(* Logix 5000 project; controller TFF vendor 1 type 14 code 107 rev 34.11; software revision 34.03; part 26 of 36 *)
(* tags used below, declared in another part *)
   Address : DINT;   // Temp Address
   Index : DINT;   // Index
   AI101 : ALIAS FOR AnalogPoint[10];   // Filtrate Conductivity
   AI102 : ALIAS FOR AnalogPoint[11];   // Filtrate UV
   AI103 : ALIAS FOR AnalogPoint[12];   // Filtrate UV
   AI104 : ALIAS FOR AnalogPoint[9];   // Filtrate pH
   AlarmControl : AlarmControl;   // Alarm Control
   CPU_Scanning : BOOL;   // System Scanning Flag
   DigitalOutput : BOOL[256];   // Digital Output Array these bits are sent to output cards.
   DigitalPoint : DigitalPoint[150];   // Digital Point Array
   Drive : Drive[11];   // Drives Array
   FI101 : ALIAS FOR AnalogPoint[2];   // Filtrate Flow
   MIX001 : ALIAS FOR AnalogPoint[14];   // Mixer Speed
   Mixer : Mixer;   // Mixer config. structure
   Options : Options;   // Options List
   Phase0 : ALIAS FOR Phase[0];   // Phase 0
   PI001 : ALIAS FOR AnalogPoint[5];   // Feed Pressure
   PI002 : ALIAS FOR AnalogPoint[6];   // Retentate Pressure
   PI101 : ALIAS FOR AnalogPoint[7];   // Filtrate Pressure
   PI401 : ALIAS FOR AnalogPoint[8];   // Transfer Pump Pressure
   PLCFault : FaultRecordType;   // PLC Major Fault Record
   Rack_Murr_Node1_TF2S : IO_Station;   // Status of Node 1 TF2S
   Rack_Murr_Node1_TF3S : IO_Station;   // Status of Node 1 TF3S
   Rack_Murr_Node4_Instrum_TFF1 : IO_Station;   // Status of Node 4 Instrum TFF1
   Rack_Murr_Node4_Instrum_TFF2 : IO_Station;   // Status of Node 4 Instrum TFF2
   Rack_Murr_Node4_Instrum_TFF3 : IO_Station;   // Status of Node 4 Instrum TFF3
   Rack_Murr_Node4_Instrum_TFF4 : IO_Station;   // Status of Node 4 Instrum TFF4
   Rack_Murr_Node4_Instrum_TFF5 : IO_Station;   // Status of Node 4 Instrum TFF5
   Rack_Murr_Node5_Tank100 : IO_Station;   // Status of Node 5 Tank 100L
   Rack_Murr_Node5_Tank250 : IO_Station;   // Status of Node 5 Tank 250L
   Rack_Murr_Node5_Tank50 : IO_Station;   // Status of Node 5 Tank 50L
   RawAnalogInputArray : INT[50];   // Array of analog input raw
   SIC003 : ALIAS FOR Drive[3];   // Mixer
   SIC003DF : ALIAS FOR DigitalPoint[14];   // Mixer Defect
   SRL001 : ALIAS FOR DigitalPoint[15];   // Tank Skid Remote / Standalone
   SysControl : SysControl;   // General system status and command
   Tank : TankManagement;   // Tank Management
   ThisSystem : SystemType;
   TI001 : ALIAS FOR AnalogPoint[13];   // Feed Bag Temperature
   WI001 : ALIAS FOR AnalogPoint[15];   // Feed Bag Weight
   YA10 : ALIAS FOR DigitalPoint[59];   // PLC Program Major Fault
(* Process, continued *)

ROUTINE Drive_SIC003_Mixer   (* ladder *)
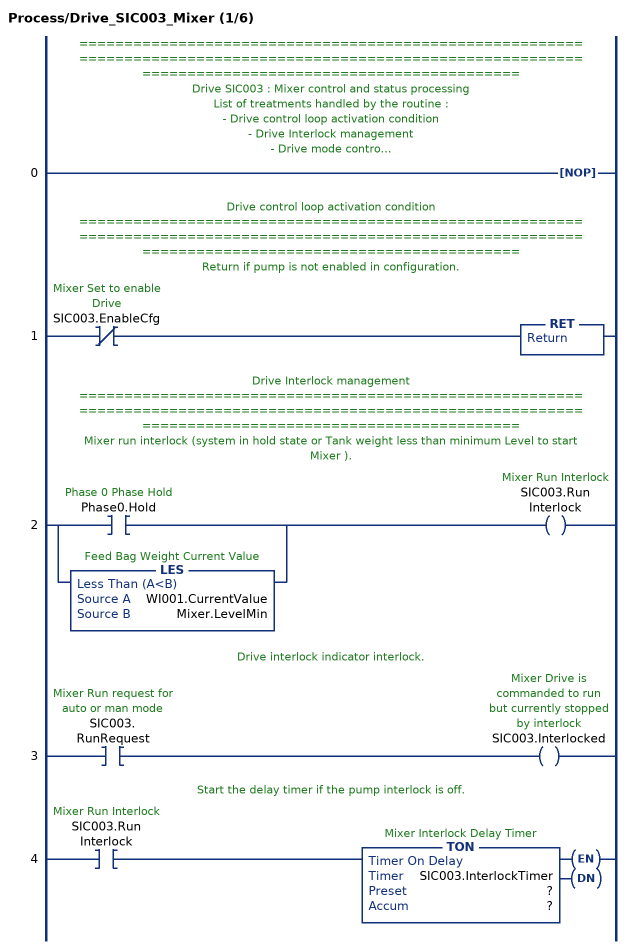
   // ==========================================================================================================================================================
   //                                                        Drive SIC003 : Mixer control and status processing
   //                                                     List of treatments handled by the routine :
   //                                                          - Drive control loop activation condition
   //                                                          - Drive Interlock management
   //                                                          - Drive mode control
   //                                                          - Drive run command control
   //                                                          - Drive status management
   //                                                          - Drive status for HMI
   //                                                          - Drive DigitalOutput control
   //                                                     -----------------------------------------------------------------------------------------------------------------------------------------------------
   //                                                     History
   //                                                          2019-AUG-13 - Actemium - B. Roch - Initial version for Candidate Release 3.00.00.00.a
   //                                                          2019-OCT-25 - Actemium - B. Roch - Modification for Candidate Release 3.00.00.00.d
   //                                                      - Add Mixer standalone condition to stop mixer
   // ==========================================================================================================================================================
   0: NOP();
   // Drive control loop activation condition
   // ==========================================================================================================================================================
   // Return if pump is not enabled in configuration.
   1: XIO(SIC003.EnableCfg)RET();
   // Drive Interlock management
   // ==========================================================================================================================================================
   // Mixer run interlock (system in hold state or Tank weight less than minimum Level to start Mixer ).
   2: [XIC(Phase0.Hold) ,LES(WI001.CurrentValue,Mixer.LevelMin) ]OTE(SIC003.RunInterlock);
   // Drive interlock indicator interlock.
   3: XIC(SIC003.RunRequest)OTE(SIC003.Interlocked);
   // Start the delay timer if the pump interlock is off.
   4: XIC(SIC003.RunInterlock)TON(SIC003.InterlockTimer,?,?);
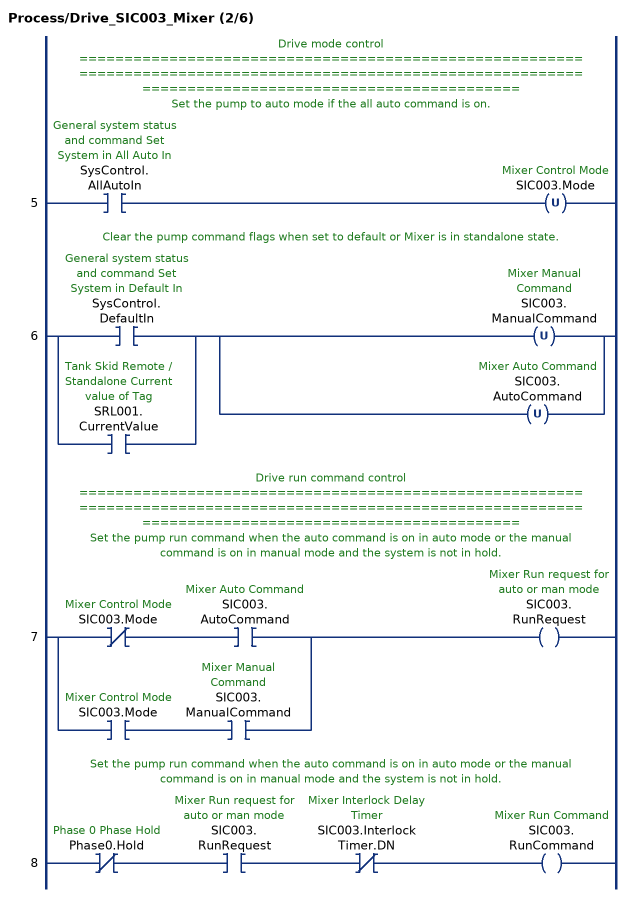
   // Drive mode control
   // ==========================================================================================================================================================
   // Set the pump to auto mode if the all auto command is on.
   5: XIC(SysControl.AllAutoIn)OTU(SIC003.Mode);
   // Clear the pump command flags when set to default or Mixer is in standalone state.
   6: [XIC(SysControl.DefaultIn) ,XIC(SRL001.CurrentValue) ][OTU(SIC003.ManualCommand) ,OTU(SIC003.AutoCommand) ];
   // Drive run command control
   // ==========================================================================================================================================================
   // Set the pump run command when the auto command is on in auto mode or the manual command is on in manual mode and the system is not in hold.
   7: [XIO(SIC003.Mode) XIC(SIC003.AutoCommand) ,XIC(SIC003.Mode) XIC(SIC003.ManualCommand) ]OTE(SIC003.RunRequest);
   // Set the pump run command when the auto command is on in auto mode or the manual command is on in manual mode and the system is not in hold.
   8: XIO(Phase0.Hold)XIC(SIC003.RunRequest)XIO(SIC003.InterlockTimer.DN)OTE(SIC003.RunCommand);
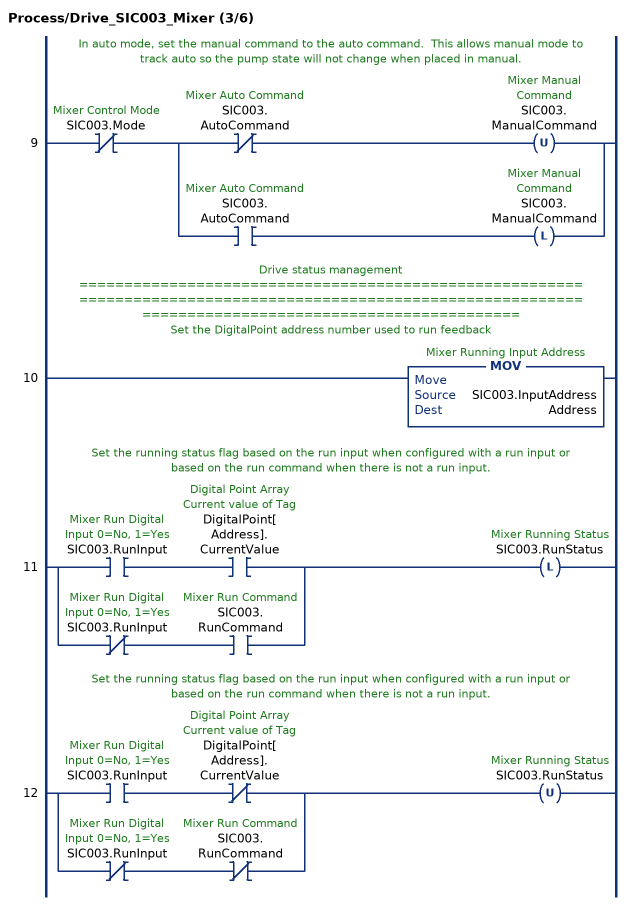
   // In auto mode, set the manual command to the auto command.  This allows manual mode to track auto so the pump state will not change when placed in manual.
   9: XIO(SIC003.Mode)[XIO(SIC003.AutoCommand) OTU(SIC003.ManualCommand) ,XIC(SIC003.AutoCommand) OTL(SIC003.ManualCommand) ];
   // Drive status management
   // ==========================================================================================================================================================
   // Set the DigitalPoint address number used to run feedback
   10: MOV(SIC003.InputAddress,Address);
   // Set the running status flag based on the run input when configured with a run input or based on the run command when there is not a run input.
   11: [XIC(SIC003.RunInput) XIC(DigitalPoint[Address].CurrentValue) ,XIO(SIC003.RunInput) XIC(SIC003.RunCommand) ]OTL(SIC003.RunStatus);
   // Set the running status flag based on the run input when configured with a run input or based on the run command when there is not a run input.
   12: [XIC(SIC003.RunInput) XIO(DigitalPoint[Address].CurrentValue) ,XIO(SIC003.RunInput) XIO(SIC003.RunCommand) ]OTU(SIC003.RunStatus);
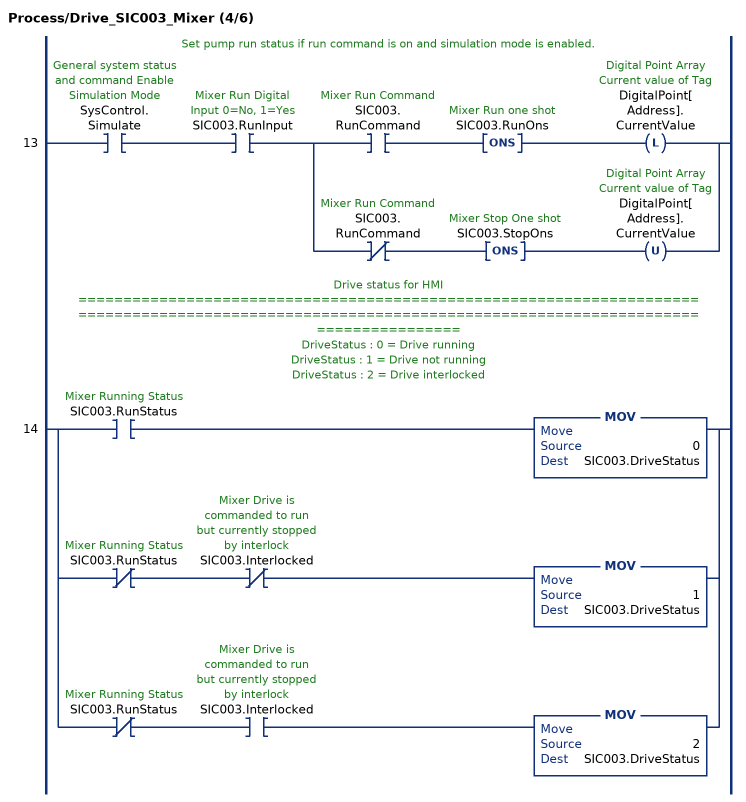
   // Set pump run status if run command is on and simulation mode is enabled.
   13: XIC(SysControl.Simulate)XIC(SIC003.RunInput)[XIC(SIC003.RunCommand) ONS(SIC003.RunOns) OTL(DigitalPoint[Address].CurrentValue) ,XIO(SIC003.RunCommand) ONS(SIC003.StopOns) OTU(DigitalPoint[Address].CurrentValue) ];
   // Drive status for HMI
   // ==========================================================================================================================================================
   //  DriveStatus : 0 = Drive running
   //  DriveStatus : 1 = Drive not running
   //  DriveStatus : 2 = Drive interlocked
   14: [XIC(SIC003.RunStatus) MOV(0,SIC003.DriveStatus) ,XIO(SIC003.RunStatus) XIO(SIC003.Interlocked) MOV(1,SIC003.DriveStatus) ,XIO(SIC003.RunStatus) XIC(SIC003.Interlocked) MOV(2,SIC003.DriveStatus) ];
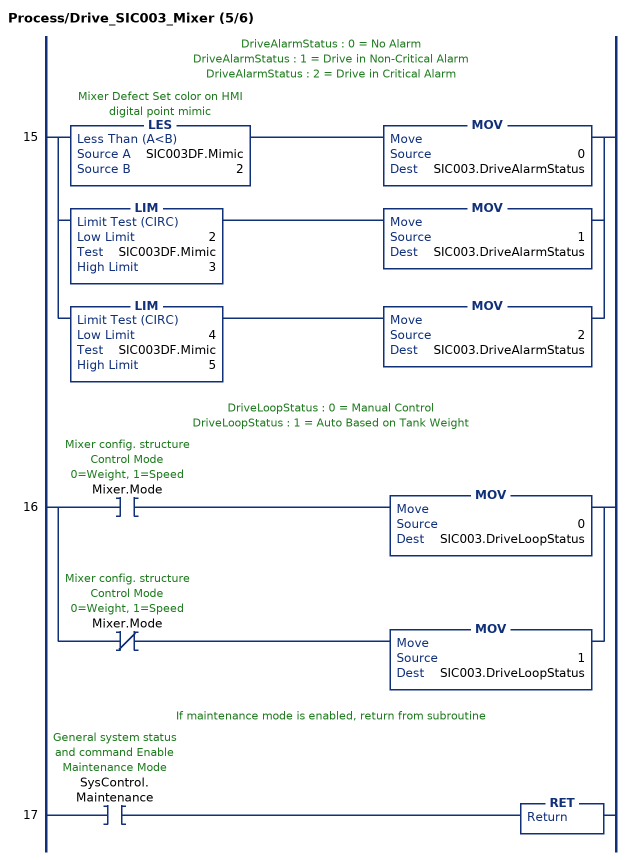
   // DriveAlarmStatus : 0 = No Alarm
   //  DriveAlarmStatus : 1 = Drive in Non-Critical Alarm
   //  DriveAlarmStatus : 2 = Drive in Critical Alarm
   15: [LES(SIC003DF.Mimic,2) MOV(0,SIC003.DriveAlarmStatus) ,LIM(2,SIC003DF.Mimic,3) MOV(1,SIC003.DriveAlarmStatus) ,LIM(4,SIC003DF.Mimic,5) MOV(2,SIC003.DriveAlarmStatus) ];
   // DriveLoopStatus : 0 = Manual Control
   //  DriveLoopStatus : 1 = Auto Based on Tank Weight
   16: [XIC(Mixer.Mode) MOV(0,SIC003.DriveLoopStatus) ,XIO(Mixer.Mode) MOV(1,SIC003.DriveLoopStatus) ];
   // If maintenance mode is enabled, return from subroutine
   17: XIC(SysControl.Maintenance)RET();
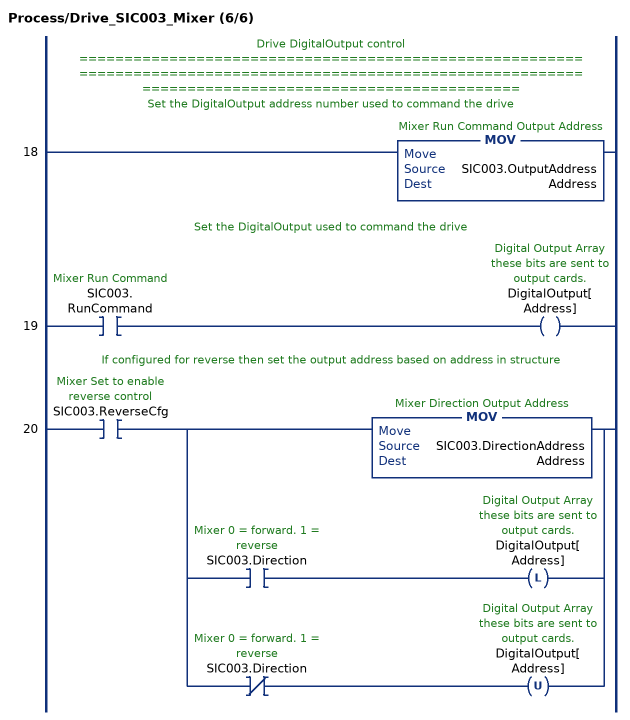
   // Drive DigitalOutput control
   // ==========================================================================================================================================================
   // Set the DigitalOutput address number used to command the drive
   18: MOV(SIC003.OutputAddress,Address);
   // Set the DigitalOutput used to command the drive
   19: XIC(SIC003.RunCommand)OTE(DigitalOutput[Address]);
   // If configured for reverse then set the output address based on address in structure
   20: XIC(SIC003.ReverseCfg)[MOV(SIC003.DirectionAddress,Address) ,XIC(SIC003.Direction) OTL(DigitalOutput[Address]) ,XIO(SIC003.Direction) OTU(DigitalOutput[Address]) ];
END_ROUTINE

ROUTINE Drives   (* ladder *)
// Pump Control Routine
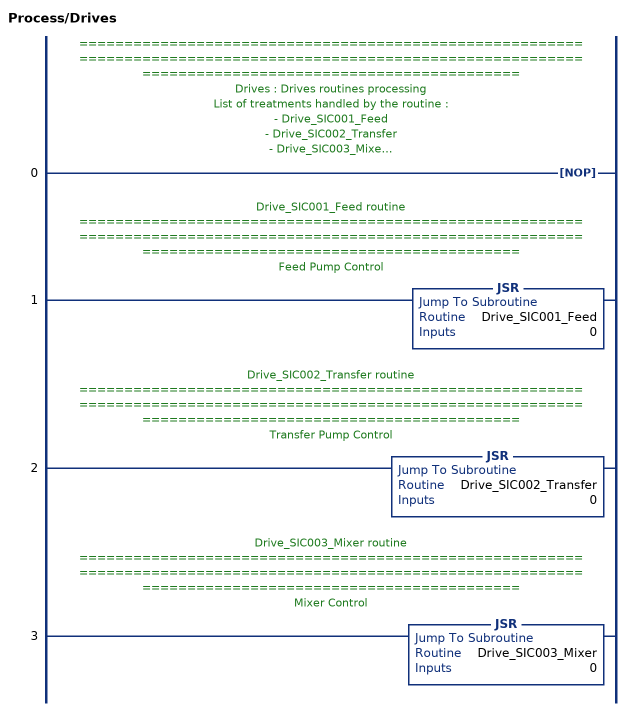
   // ==========================================================================================================================================================
   //                                                                                                                           Drives : Drives routines processing
   //                                                     List of treatments handled by the routine :
   //                                                          - Drive_SIC001_Feed
   //                                                          - Drive_SIC002_Transfer
   //                                                          - Drive_SIC003_Mixer
   //                                                     -----------------------------------------------------------------------------------------------------------------------------------------------------
   //                                                     History
   //                                                         2019-AUG-13 - Actemium - B. Roch - Initial version for Candidate Release 3.00.00.00.a
   // ==========================================================================================================================================================
   0: NOP();
   // Drive_SIC001_Feed routine
   // ==========================================================================================================================================================
   // Feed Pump Control
   1: JSR(Drive_SIC001_Feed,0);
   // Drive_SIC002_Transfer routine
   // ==========================================================================================================================================================
   // Transfer Pump Control
   2: JSR(Drive_SIC002_Transfer,0);
   // Drive_SIC003_Mixer routine
   // ==========================================================================================================================================================
   // Mixer Control
   3: JSR(Drive_SIC003_Mixer,0);
END_ROUTINE

ROUTINE FaultRoutine   (* ladder *)
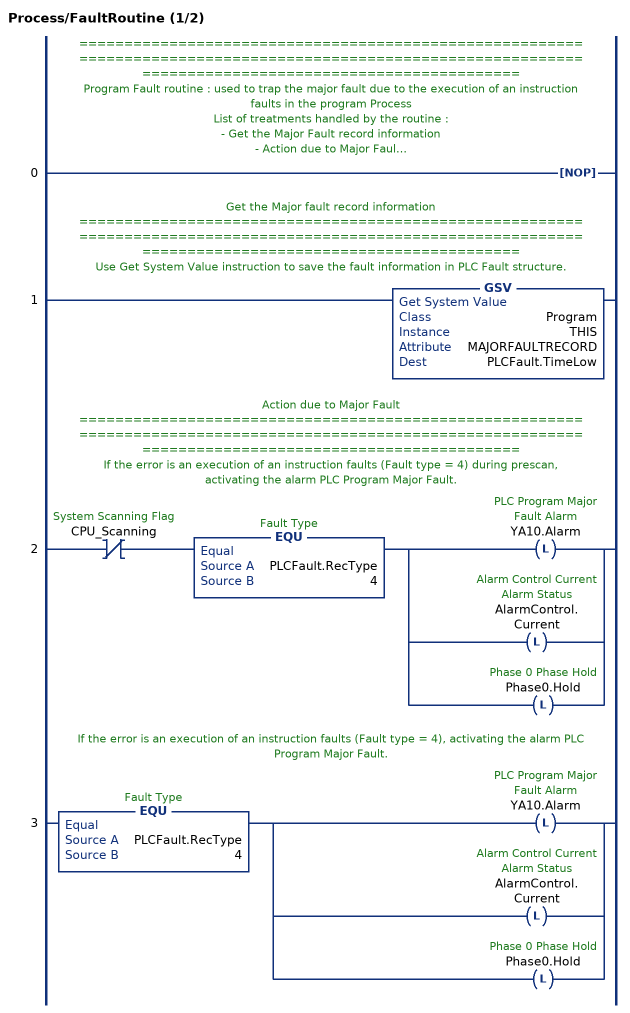
   // ==========================================================================================================================================================
   //                                                               Program Fault routine : used to trap the major fault due to the execution of an instruction faults in the program Process
   //                                                     List of treatments handled by the routine :
   //                                                          - Get the Major Fault record information
   //                                                          - Action due to Major Fault
   //                                                     -----------------------------------------------------------------------------------------------------------------------------------------------------
   //                                                     History
   //                                                          2019-AUG-13 - Actemium - B. Roch - Initial version for Candidate Release 3.00.00.00.a
   // ==========================================================================================================================================================
   0: NOP();
   // Get the Major fault record information
   // ==========================================================================================================================================================
   // Use Get System Value instruction to save the fault information in PLC Fault structure.
   1: GSV(Program,THIS,MAJORFAULTRECORD,PLCFault.TimeLow);
   // Action due to Major Fault
   // ==========================================================================================================================================================
   // If the error is an execution of an instruction faults (Fault type = 4) during prescan, activating the alarm PLC Program Major Fault.
   2: XIO(CPU_Scanning)EQU(PLCFault.RecType,4)[OTL(YA10.Alarm) ,OTL(AlarmControl.Current) ,OTL(Phase0.Hold) ];
   // If the error is an execution of an instruction faults (Fault type = 4), activating the alarm PLC Program Major Fault.
   3: EQU(PLCFault.RecType,4)[OTL(YA10.Alarm) ,OTL(AlarmControl.Current) ,OTL(Phase0.Hold) ];
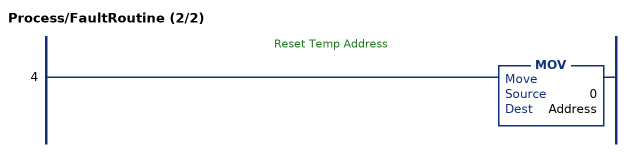
   // Reset Temp Address
   4: MOV(0,Address);
END_ROUTINE

ROUTINE InputAnalogPoint   (* ladder *)
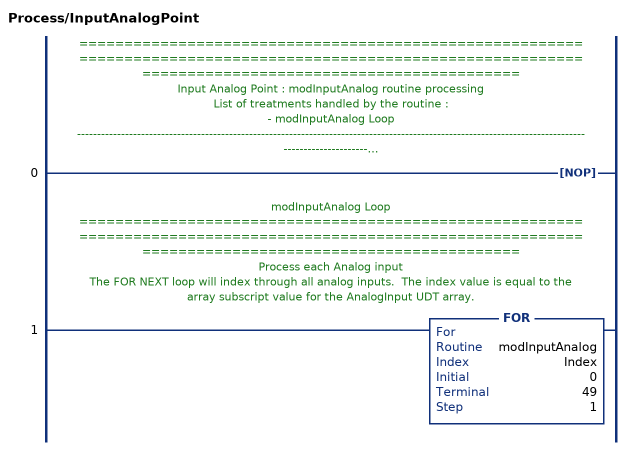
   // ==========================================================================================================================================================
   //                                                                                                             Input Analog Point : modInputAnalog routine processing
   //                                                     List of treatments handled by the routine :
   //                                                          - modInputAnalog Loop
   //                                                     -----------------------------------------------------------------------------------------------------------------------------------------------------
   //                                                     History
   //                                                          2019-AUG-13 - Actemium - B. Roch - Initial version for Candidate Release 3.00.00.00.a
   // ==========================================================================================================================================================
   0: NOP();
   // modInputAnalog Loop
   // ==========================================================================================================================================================
   // Process each Analog input
   // The FOR NEXT loop will index through all analog inputs.  The index value is equal to the array subscript value for the AnalogInput UDT array.
   1: FOR(modInputAnalog,Index,0,49,1);
END_ROUTINE

ROUTINE InputAnalogRaw   (* ladder *)
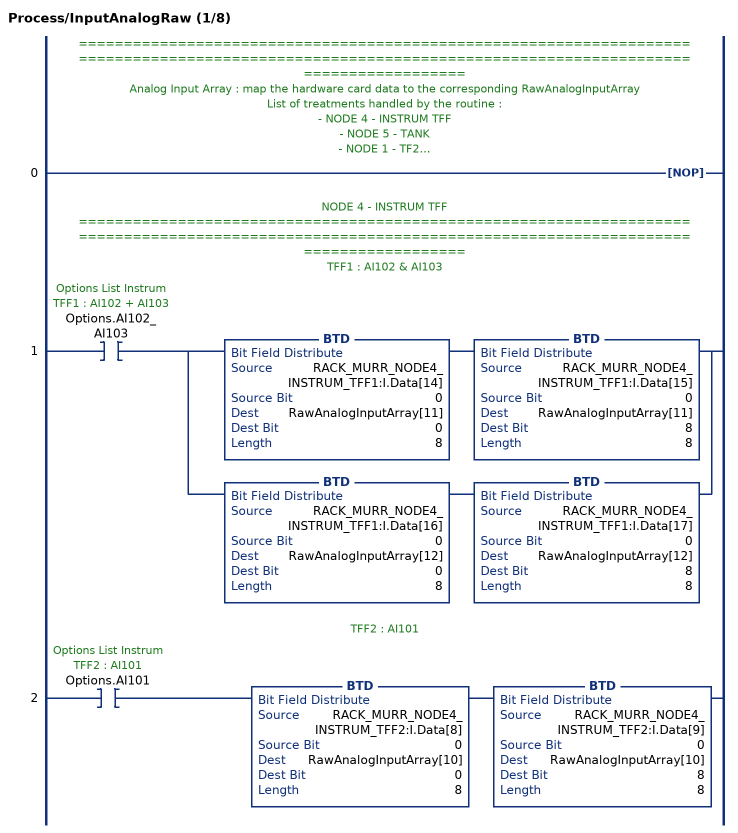
   // ==========================================================================================================================================================
   //                                                                                          Analog Input Array : map the hardware card data to the corresponding RawAnalogInputArray
   //                                                     List of treatments handled by the routine :
   //                                                     - NODE 4 - INSTRUM TFF
   //                                                     - NODE 5 - TANK
   //                                                     - NODE 1 - TF2S
   //                                                     - NODE 1 - TF3S
   //                                                     -----------------------------------------------------------------------------------------------------------------------------------------------------
   //                                                     History
   //                                                          2019-AUG-13 - Actemium - B. Roch - Initial version for Candidate Release 3.00.00.00.a
   // ==========================================================================================================================================================
   0: NOP();
   // NODE 4 - INSTRUM TFF
   // ==========================================================================================================================================================
   // TFF1 : AI102 & AI103
   1: XIC(Options.AI102_AI103)[BTD(RACK_MURR_NODE4_INSTRUM_TFF1:I.Data[14],0,RawAnalogInputArray[11],0,8) BTD(RACK_MURR_NODE4_INSTRUM_TFF1:I.Data[15],0,RawAnalogInputArray[11],8,8) ,BTD(RACK_MURR_NODE4_INSTRUM_TFF1:I.Data[16],0,RawAnalogInputArray[12],0,8) BTD(RACK_MURR_NODE4_INSTRUM_TFF1:I.Data[17],0,RawAnalogInputArray[12],8,8) ];
   // TFF2 : AI101
   2: XIC(Options.AI101)BTD(RACK_MURR_NODE4_INSTRUM_TFF2:I.Data[8],0,RawAnalogInputArray[10],0,8)BTD(RACK_MURR_NODE4_INSTRUM_TFF2:I.Data[9],0,RawAnalogInputArray[10],8,8);
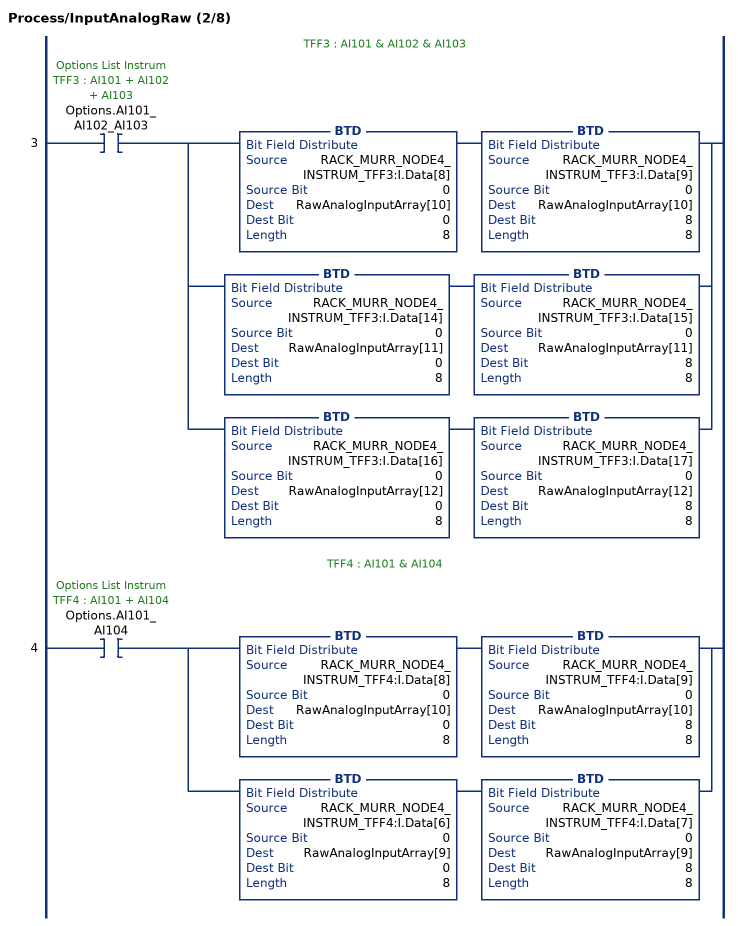
   // TFF3 : AI101 & AI102 & AI103
   3: XIC(Options.AI101_AI102_AI103)[BTD(RACK_MURR_NODE4_INSTRUM_TFF3:I.Data[8],0,RawAnalogInputArray[10],0,8) BTD(RACK_MURR_NODE4_INSTRUM_TFF3:I.Data[9],0,RawAnalogInputArray[10],8,8) ,BTD(RACK_MURR_NODE4_INSTRUM_TFF3:I.Data[14],0,RawAnalogInputArray[11],0,8) BTD(RACK_MURR_NODE4_INSTRUM_TFF3:I.Data[15],0,RawAnalogInputArray[11],8,8) ,BTD(RACK_MURR_NODE4_INSTRUM_TFF3:I.Data[16],0,RawAnalogInputArray[12],0,8) BTD(RACK_MURR_NODE4_INSTRUM_TFF3:I.Data[17],0,RawAnalogInputArray[12],8,8) ];
   // TFF4 : AI101 & AI104
   4: XIC(Options.AI101_AI104)[BTD(RACK_MURR_NODE4_INSTRUM_TFF4:I.Data[8],0,RawAnalogInputArray[10],0,8) BTD(RACK_MURR_NODE4_INSTRUM_TFF4:I.Data[9],0,RawAnalogInputArray[10],8,8) ,BTD(RACK_MURR_NODE4_INSTRUM_TFF4:I.Data[6],0,RawAnalogInputArray[9],0,8) BTD(RACK_MURR_NODE4_INSTRUM_TFF4:I.Data[7],0,RawAnalogInputArray[9],8,8) ];
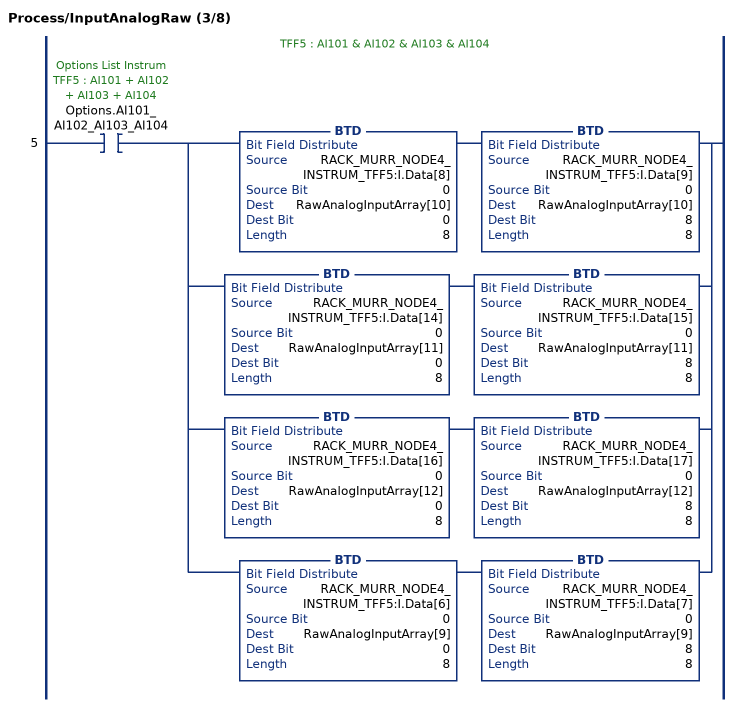
   // TFF5 : AI101 & AI102 & AI103 & AI104
   5: XIC(Options.AI101_AI102_AI103_AI104)[BTD(RACK_MURR_NODE4_INSTRUM_TFF5:I.Data[8],0,RawAnalogInputArray[10],0,8) BTD(RACK_MURR_NODE4_INSTRUM_TFF5:I.Data[9],0,RawAnalogInputArray[10],8,8) ,BTD(RACK_MURR_NODE4_INSTRUM_TFF5:I.Data[14],0,RawAnalogInputArray[11],0,8) BTD(RACK_MURR_NODE4_INSTRUM_TFF5:I.Data[15],0,RawAnalogInputArray[11],8,8) ,BTD(RACK_MURR_NODE4_INSTRUM_TFF5:I.Data[16],0,RawAnalogInputArray[12],0,8) BTD(RACK_MURR_NODE4_INSTRUM_TFF5:I.Data[17],0,RawAnalogInputArray[12],8,8) ,BTD(RACK_MURR_NODE4_INSTRUM_TFF5:I.Data[6],0,RawAnalogInputArray[9],0,8) BTD(RACK_MURR_NODE4_INSTRUM_TFF5:I.Data[7],0,RawAnalogInputArray[9],8,8) ];
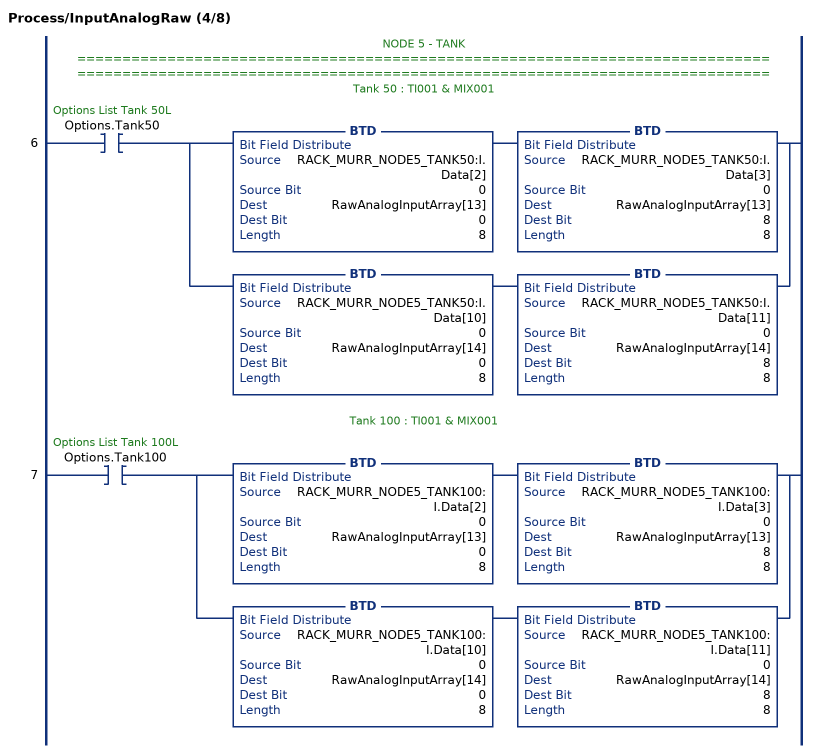
   // NODE 5 - TANK
   // ==========================================================================================================================================================
   // Tank 50 : TI001 & MIX001
   6: XIC(Options.Tank50)[BTD(RACK_MURR_NODE5_TANK50:I.Data[2],0,RawAnalogInputArray[13],0,8) BTD(RACK_MURR_NODE5_TANK50:I.Data[3],0,RawAnalogInputArray[13],8,8) ,BTD(RACK_MURR_NODE5_TANK50:I.Data[10],0,RawAnalogInputArray[14],0,8) BTD(RACK_MURR_NODE5_TANK50:I.Data[11],0,RawAnalogInputArray[14],8,8) ];
   // Tank 100 : TI001 & MIX001
   7: XIC(Options.Tank100)[BTD(RACK_MURR_NODE5_TANK100:I.Data[2],0,RawAnalogInputArray[13],0,8) BTD(RACK_MURR_NODE5_TANK100:I.Data[3],0,RawAnalogInputArray[13],8,8) ,BTD(RACK_MURR_NODE5_TANK100:I.Data[10],0,RawAnalogInputArray[14],0,8) BTD(RACK_MURR_NODE5_TANK100:I.Data[11],0,RawAnalogInputArray[14],8,8) ];
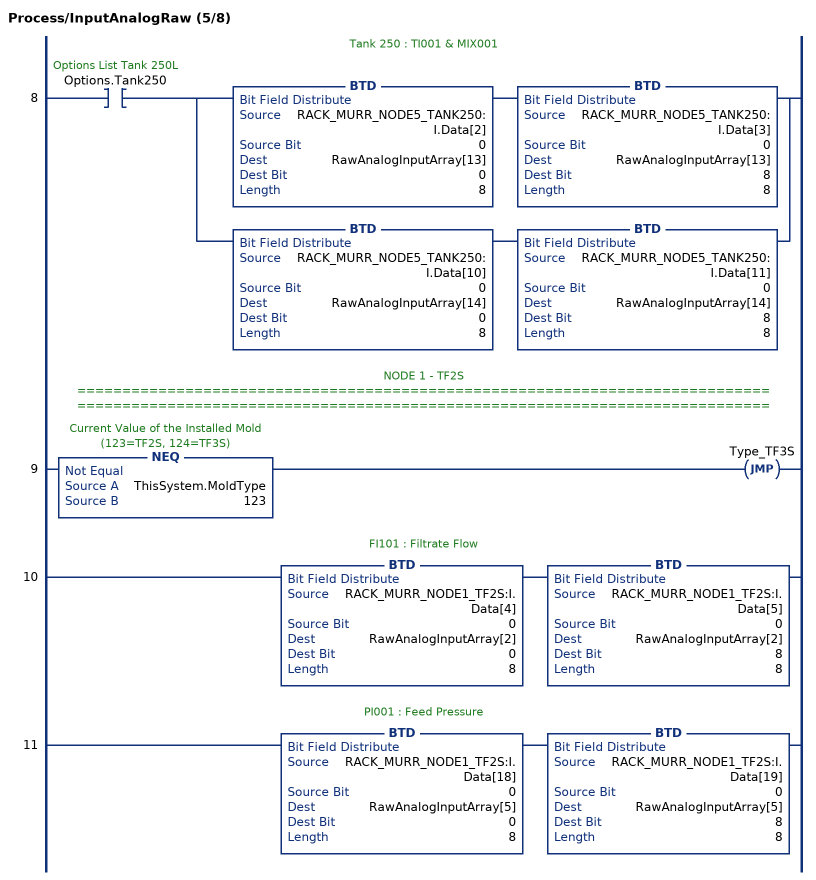
   // Tank 250 : TI001 & MIX001
   8: XIC(Options.Tank250)[BTD(RACK_MURR_NODE5_TANK250:I.Data[2],0,RawAnalogInputArray[13],0,8) BTD(RACK_MURR_NODE5_TANK250:I.Data[3],0,RawAnalogInputArray[13],8,8) ,BTD(RACK_MURR_NODE5_TANK250:I.Data[10],0,RawAnalogInputArray[14],0,8) BTD(RACK_MURR_NODE5_TANK250:I.Data[11],0,RawAnalogInputArray[14],8,8) ];
   // NODE 1 - TF2S
   // ==========================================================================================================================================================
   9: NEQ(ThisSystem.MoldType,123)JMP(Type_TF3S);
   // FI101 : Filtrate Flow
   10: BTD(RACK_MURR_NODE1_TF2S:I.Data[4],0,RawAnalogInputArray[2],0,8)BTD(RACK_MURR_NODE1_TF2S:I.Data[5],0,RawAnalogInputArray[2],8,8);
   // PI001 : Feed Pressure
   11: BTD(RACK_MURR_NODE1_TF2S:I.Data[18],0,RawAnalogInputArray[5],0,8)BTD(RACK_MURR_NODE1_TF2S:I.Data[19],0,RawAnalogInputArray[5],8,8);
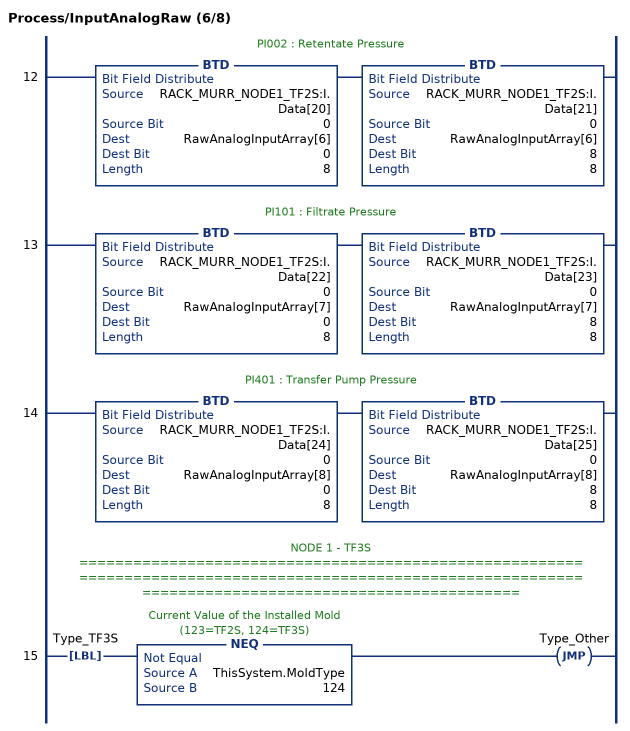
   // PI002 : Retentate Pressure
   12: BTD(RACK_MURR_NODE1_TF2S:I.Data[20],0,RawAnalogInputArray[6],0,8)BTD(RACK_MURR_NODE1_TF2S:I.Data[21],0,RawAnalogInputArray[6],8,8);
   // PI101 : Filtrate Pressure
   13: BTD(RACK_MURR_NODE1_TF2S:I.Data[22],0,RawAnalogInputArray[7],0,8)BTD(RACK_MURR_NODE1_TF2S:I.Data[23],0,RawAnalogInputArray[7],8,8);
   // PI401 : Transfer Pump Pressure
   14: BTD(RACK_MURR_NODE1_TF2S:I.Data[24],0,RawAnalogInputArray[8],0,8)BTD(RACK_MURR_NODE1_TF2S:I.Data[25],0,RawAnalogInputArray[8],8,8);
   // NODE 1 - TF3S
   // ==========================================================================================================================================================
   15: LBL(Type_TF3S)NEQ(ThisSystem.MoldType,124)JMP(Type_Other);
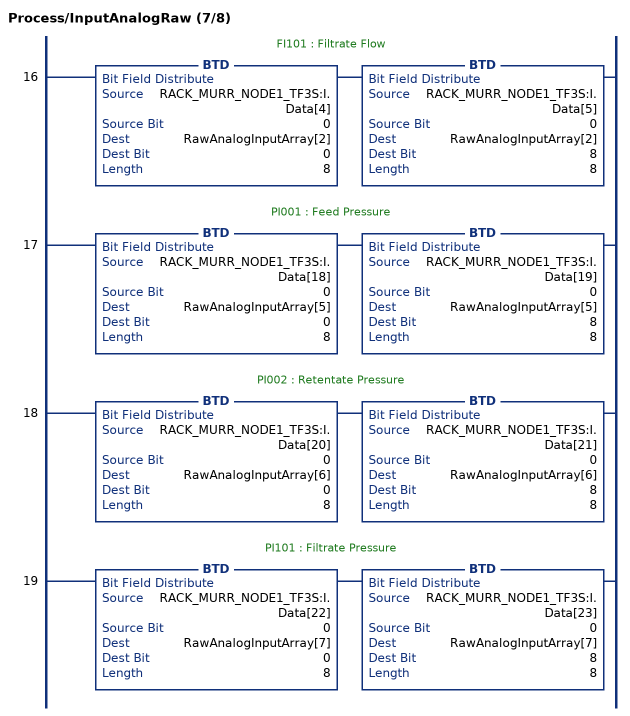
   // FI101 : Filtrate Flow
   16: BTD(RACK_MURR_NODE1_TF3S:I.Data[4],0,RawAnalogInputArray[2],0,8)BTD(RACK_MURR_NODE1_TF3S:I.Data[5],0,RawAnalogInputArray[2],8,8);
   // PI001 : Feed Pressure
   17: BTD(RACK_MURR_NODE1_TF3S:I.Data[18],0,RawAnalogInputArray[5],0,8)BTD(RACK_MURR_NODE1_TF3S:I.Data[19],0,RawAnalogInputArray[5],8,8);
   // PI002 : Retentate Pressure
   18: BTD(RACK_MURR_NODE1_TF3S:I.Data[20],0,RawAnalogInputArray[6],0,8)BTD(RACK_MURR_NODE1_TF3S:I.Data[21],0,RawAnalogInputArray[6],8,8);
   // PI101 : Filtrate Pressure
   19: BTD(RACK_MURR_NODE1_TF3S:I.Data[22],0,RawAnalogInputArray[7],0,8)BTD(RACK_MURR_NODE1_TF3S:I.Data[23],0,RawAnalogInputArray[7],8,8);
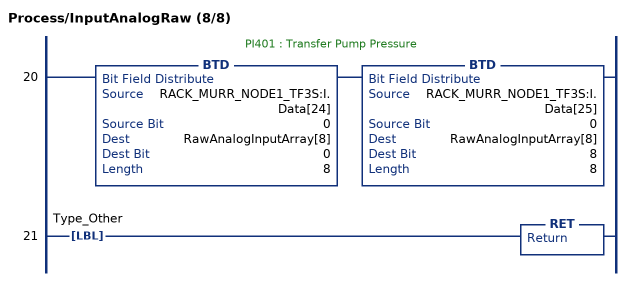
   // PI401 : Transfer Pump Pressure
   20: BTD(RACK_MURR_NODE1_TF3S:I.Data[24],0,RawAnalogInputArray[8],0,8)BTD(RACK_MURR_NODE1_TF3S:I.Data[25],0,RawAnalogInputArray[8],8,8);
   21: LBL(Type_Other)RET();
END_ROUTINE
